(* IEC 61131-3 sources: kns-port-domestic/targets/astra/src/POUs/Regul/PRG_ModbusMap_Regul, 2 files *)

(* ---- PRG_ModbusMap_Regul.decl.st ---- *)
// Назначение: слой Modbus RTU сборки для ПЛК REGUL: массивы WORD каналов устройств Modbus Serial Outer
//             Slave ↔ регистры GVL_IO (ПЧ Н1…Н3 на RS485-1, TT403 на RS485-2) и признаки обмена
//             GVL_IO.xMbOk_* по статусу каналов чтения. Заменяет мастер Modbus CODESYS с диагностикой слейвов
//             (у флагмана — слой Modbus сборки ПЛК210). Вызывается первой в MainTask только в сборке для ПЛК
//             (GVL_Const.SIM_ALLOWED = FALSE) и на стенде с Modbus TCP вместо RTU; в имитации регистры GVL_IO
//             пишет модель объекта, программа сразу выходит.
// Автор:      kr0nsch
// Версия:     0.1.0
// Документ:   targets/astra/README.md; docs/migration_checklist.md, раздел 4
// PORT: [comm] новый объект: Modbus RTU на REGUL — каналы Modbus Serial Outer Slave [F57, F58]
PROGRAM PRG_ModbusMap_Regul
VAR
    // Data каналов — привязать в «Соотнесении входов/выходов» каналов слейвов (E1, E2)
    awP101Rd : ARRAY[0..GVL_ConstRegul.MB_VFD_RD_LAST] OF WORD;  // слейв 1: канал FC3 4x 100, 4 регистра, Timer
    awP102Rd : ARRAY[0..GVL_ConstRegul.MB_VFD_RD_LAST] OF WORD;  // слейв 2: то же
    awP103Rd : ARRAY[0..GVL_ConstRegul.MB_VFD_RD_LAST] OF WORD;  // слейв 3: то же
    awP101Wr : ARRAY[0..GVL_ConstRegul.MB_VFD_WR_LAST] OF WORD;  // слейв 1: канал FC16 4x 0, 2 регистра, Timer
    awP102Wr : ARRAY[0..GVL_ConstRegul.MB_VFD_WR_LAST] OF WORD;  // слейв 2: то же
    awP103Wr : ARRAY[0..GVL_ConstRegul.MB_VFD_WR_LAST] OF WORD;  // слейв 3: то же
    awTT403Rd : ARRAY[0..GVL_ConstRegul.MB_REAL_LAST] OF WORD;   // RS485-2, слейв 10: канал FC4 3x 0, 2 регистра
    // Status каналов чтения — привязать к Status тех же каналов
    // PORT: [comm] BUILD_ERRORS 1.1: ChannelStatus — в пространстве имён PsIoDrvModbusSerialMaster
    // (имя библиотеки драйвера; PsModbusSerialMaster из DPA-302.1 в Astra.IDE 1.7.2.2 не находится — C0077)
    // PORT: [comm] проверить в Astra.IDE — привязка Status каналов к этим переменным [F58] (E2)
    eP101Status : PsIoDrvModbusSerialMaster.ChannelStatus;
    eP102Status : PsIoDrvModbusSerialMaster.ChannelStatus;
    eP103Status : PsIoDrvModbusSerialMaster.ChannelStatus;
    eTT403Status : PsIoDrvModbusSerialMaster.ChannelStatus;
    uTT403 : PL.U_RealBits;     // REAL из двух регистров
END_VAR

(* ---- PRG_ModbusMap_Regul.impl.st ---- *)
// В имитации регистры и признаки обмена GVL_IO пишет модель объекта (PRG_PlantModel)
IF GVL_Sim.xSimulation THEN
    RETURN;
END_IF

// 1. ПЧ Н1…Н3, чтение: слово состояния, фактическая частота, ток, код аварии (те же регистры, что у мастера CODESYS)
GVL_IO.wP101_STW := awP101Rd[GVL_ConstRegul.MB_VFD_RD_STW];
GVL_IO.uiP101_FACT := WORD_TO_UINT(awP101Rd[GVL_ConstRegul.MB_VFD_RD_FACT]);
GVL_IO.uiIT111 := WORD_TO_UINT(awP101Rd[GVL_ConstRegul.MB_VFD_RD_IT]);
GVL_IO.uiP101_FCODE := WORD_TO_UINT(awP101Rd[GVL_ConstRegul.MB_VFD_RD_FCODE]);

GVL_IO.wP102_STW := awP102Rd[GVL_ConstRegul.MB_VFD_RD_STW];
GVL_IO.uiP102_FACT := WORD_TO_UINT(awP102Rd[GVL_ConstRegul.MB_VFD_RD_FACT]);
GVL_IO.uiIT121 := WORD_TO_UINT(awP102Rd[GVL_ConstRegul.MB_VFD_RD_IT]);
GVL_IO.uiP102_FCODE := WORD_TO_UINT(awP102Rd[GVL_ConstRegul.MB_VFD_RD_FCODE]);

GVL_IO.wP103_STW := awP103Rd[GVL_ConstRegul.MB_VFD_RD_STW];
GVL_IO.uiP103_FACT := WORD_TO_UINT(awP103Rd[GVL_ConstRegul.MB_VFD_RD_FACT]);
GVL_IO.uiIT131 := WORD_TO_UINT(awP103Rd[GVL_ConstRegul.MB_VFD_RD_IT]);
GVL_IO.uiP103_FCODE := WORD_TO_UINT(awP103Rd[GVL_ConstRegul.MB_VFD_RD_FCODE]);

// 2. ПЧ Н1…Н3, запись: слово управления и задание частоты. PRG_FieldOut пишет их в конце MainTask, поэтому
//    в канал уходят значения прошлого цикла (20 мс — меньше периода опроса)
awP101Wr[GVL_ConstRegul.MB_VFD_WR_CTW] := GVL_IO.wP101_CTW;
awP101Wr[GVL_ConstRegul.MB_VFD_WR_FREF] := UINT_TO_WORD(GVL_IO.uiP101_FREF);
awP102Wr[GVL_ConstRegul.MB_VFD_WR_CTW] := GVL_IO.wP102_CTW;
awP102Wr[GVL_ConstRegul.MB_VFD_WR_FREF] := UINT_TO_WORD(GVL_IO.uiP102_FREF);
awP103Wr[GVL_ConstRegul.MB_VFD_WR_CTW] := GVL_IO.wP103_CTW;
awP103Wr[GVL_ConstRegul.MB_VFD_WR_FREF] := UINT_TO_WORD(GVL_IO.uiP103_FREF);

// 3. TT403: REAL из двух регистров, старшее слово первым (HL). Неконечное значение (NaN, ±Inf)
//    PL.FB_AnalogInput считает недостоверным (ClassifySignal)
uTT403.dwValue := SHL(WORD_TO_DWORD(awTT403Rd[GVL_ConstRegul.MB_REAL_HI]), GVL_ConstRegul.MB_WORD_BITS)
                  OR WORD_TO_DWORD(awTT403Rd[GVL_ConstRegul.MB_REAL_LO]);
GVL_IO.rTT403 := uTT403.rValue;

// 4. Признаки обмена — по статусу каналов чтения (запись идёт тем же слейвам по той же линии)
GVL_IO.xMbOk_RS485_1_S1 := F_MbStatusOk_Regul(iStatus := TO_INT(eP101Status));
GVL_IO.xMbOk_RS485_1_S2 := F_MbStatusOk_Regul(iStatus := TO_INT(eP102Status));
GVL_IO.xMbOk_RS485_1_S3 := F_MbStatusOk_Regul(iStatus := TO_INT(eP103Status));
GVL_IO.xMbOk_RS485_2_S10 := F_MbStatusOk_Regul(iStatus := TO_INT(eTT403Status));
